FUNCTION_BLOCK pusher_position (* Basic Function Block Type *)
  (* Standard: 61499-2 *)
  (* Version 0.0, 10/22/2026, macie, Schneider Electric, Template *)
  PACKAGE Main;
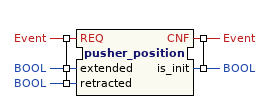
  EVENT_INPUT
    REQ WITH extended, retracted; (* Normal Execution Request *)
  END_EVENT
  EVENT_OUTPUT
    CNF WITH is_init; (* Execution Confirmation *)
  END_EVENT
  VAR_INPUT
    extended : BOOL; (* Input event qualifier *)
    retracted : BOOL;
  END_VAR
  VAR_OUTPUT
    is_init : BOOL;
  END_VAR
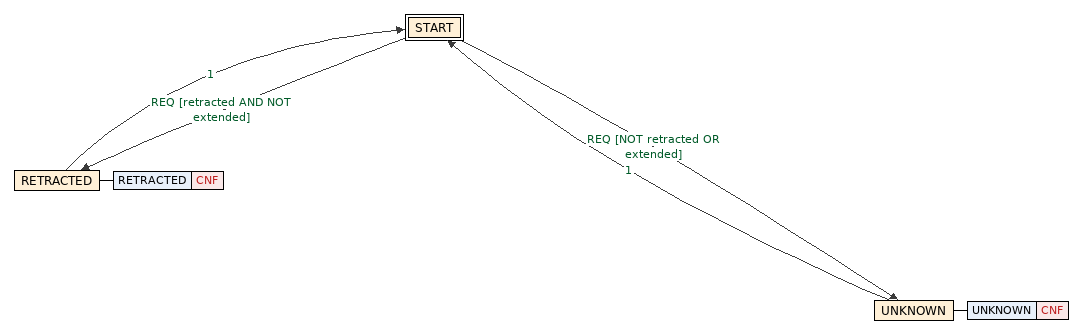
  EC_STATES
    START; (* Initial State *)
    RETRACTED : RETRACTED -> CNF; (* Normal execution *)
    UNKNOWN : UNKNOWN -> CNF;
  END_STATES
  EC_TRANSITIONS
    START TO RETRACTED := REQ [retracted AND NOT extended];
    RETRACTED TO START := 1;
    START TO UNKNOWN := REQ [NOT retracted OR extended];
    UNKNOWN TO START := 1;
  END_TRANSITIONS
  ALGORITHM RETRACTED IN ST: (* Initialization algorithm *)
;
is_init := TRUE;
  END_ALGORITHM
  ALGORITHM UNKNOWN IN ST:
;
is_init := FALSE;
  END_ALGORITHM
END_FUNCTION_BLOCK
